FUNCTION_BLOCK FB_Tank_Target EXTENDS FB_SFC_Cycle IMPLEMENTS ITF_FB_SFC_Cycle
VAR_INPUT
	//eElementID			: E_Element_List;
	valOutlet		: E_Pis_Name;
	valLine			: E_Pis_Name;
	valTriBlender	: E_Pis_Name;
	valDrain		: E_Pis_Name;	
	valCIP			: E_Pis_Name;	
END_VAR
VAR_OUTPUT
END_VAR
VAR
	//refElement		: REFERENCE TO FB_Element;
	//refState_Long		: REFERENCE TO E_Element_State_Long;
	eReq				: E_Tank_Target;
	eProcess			: E_Tank_Target;
	eStatus				: E_Tank_Target;
	
	fbPis				: FB_Piston;
	stPis_Outlet		: REFERENCE TO ST_Piston;
	stPis_Line			: REFERENCE TO ST_Piston;
	stPis_TriBlender	: REFERENCE TO ST_Piston;
	stPis_Drain			: REFERENCE TO ST_Piston;
	stPis_CIP			: REFERENCE TO ST_Piston;

	tonDrainTime: TON;
	rt_Req_Reset: R_TRIG;
	stTankLevel			:	ST_Tank_Level	;
END_VAR
VAR_IN_OUT


END_VAR

act_GetReference();

act_Oper();
IF NOT Init.x THEN;
	act_Status();
END_IF

tonDrainTime(PT:=T#1M, 
	IN:=(eStatus=E_Tank_Target.eDrain AND stTankLevel.e_state=E_Tank_Level.eEmpty)
			OR 
		eStatus=E_Tank_Target.eClose_DrainPipe);
IF tonDrainTime.Q 
AND eReq=E_Tank_Target.eNone
AND eProcess=E_Tank_Target.eNone
THEN;
	eReq:=E_Tank_Target.eClose;
END_IF

m_Request_Reset(memo:=rt_Req_Reset);//

ACTION _aCIP_active:
bStepDone:=FALSE;
IF TRUE 
AND eStatus=E_Tank_Target.eCIP
THEN;
	bStepDone:=TRUE;
END_IF
END_ACTION

ACTION _aCIP_entry:
fbPis.m_SetByRecipe(stPis:=stPis_Outlet, 		req:=E_Piston_Recipe_State.Act);
fbPis.m_SetByRecipe(stPis:=stPis_Line, 		req:=E_Piston_Recipe_State.Release);
fbPis.m_SetByRecipe(stPis:=stPis_TriBlender, 	req:=E_Piston_Recipe_State.Release);
fbPis.m_SetByRecipe(stPis:=stPis_Drain, 		req:=E_Piston_Recipe_State.Act);
fbPis.m_SetByRecipe(stPis:=stPis_CIP, 			req:=E_Piston_Recipe_State.Act);
END_ACTION

ACTION _aClose_active:
bStepDone:=FALSE;
IF TRUE 
AND eStatus=E_Tank_Target.eClose
THEN;
	bStepDone:=TRUE;
END_IF
END_ACTION

ACTION _aClose_entry:
fbPis.m_SetByRecipe(stPis:=stPis_Outlet, 		req:=E_Piston_Recipe_State.Release);
fbPis.m_SetByRecipe(stPis:=stPis_Line, 			req:=E_Piston_Recipe_State.Release);
fbPis.m_SetByRecipe(stPis:=stPis_TriBlender, 	req:=E_Piston_Recipe_State.Release);
fbPis.m_SetByRecipe(stPis:=stPis_Drain, 		req:=E_Piston_Recipe_State.Release);
fbPis.m_SetByRecipe(stPis:=stPis_CIP, 			req:=E_Piston_Recipe_State.Release);
END_ACTION

ACTION _aDone_entry:
eProcess:=E_Tank_Target.eNone;
eReq:=E_Tank_Target.eNone;
eStatus:=E_Tank_Target.eNone;
bRun:=FALSE;
bDone:=TRUE;
END_ACTION

ACTION _aDrain_active:
bStepDone:=FALSE;
IF TRUE 
AND eStatus=E_Tank_Target.eDrain
THEN;
	bStepDone:=TRUE;
END_IF
END_ACTION

ACTION _aDrain_entry:
fbPis.m_SetByRecipe(stPis:=stPis_Outlet, 		req:=E_Piston_Recipe_State.Act);
fbPis.m_SetByRecipe(stPis:=stPis_Line, 			req:=E_Piston_Recipe_State.Release);
fbPis.m_SetByRecipe(stPis:=stPis_TriBlender, 	req:=E_Piston_Recipe_State.Release);
fbPis.m_SetByRecipe(stPis:=stPis_Drain, 		req:=E_Piston_Recipe_State.Act);
fbPis.m_SetByRecipe(stPis:=stPis_CIP, 			req:=E_Piston_Recipe_State.Release);
END_ACTION

ACTION _aDrainPipe_active:
bStepDone:=FALSE;
IF TRUE 
AND eStatus=E_Tank_Target.eClose_DrainPipe
THEN;
	bStepDone:=TRUE;
END_IF
END_ACTION

ACTION _aDrainPipe_entry:
fbPis.m_SetByRecipe(stPis:=stPis_Outlet, 		req:=E_Piston_Recipe_State.Release);
fbPis.m_SetByRecipe(stPis:=stPis_Line, 			req:=E_Piston_Recipe_State.Release);
fbPis.m_SetByRecipe(stPis:=stPis_TriBlender, 	req:=E_Piston_Recipe_State.Release);
fbPis.m_SetByRecipe(stPis:=stPis_Drain, 		req:=E_Piston_Recipe_State.Act);
fbPis.m_SetByRecipe(stPis:=stPis_CIP, 			req:=E_Piston_Recipe_State.Release);
END_ACTION

ACTION _aInit_active:
SFCReset:=FALSE;
END_ACTION

ACTION _aInit_exit:
eProcess:=E_Tank_Target.eNone;
eReq:=E_Tank_Target.eNone;
END_ACTION

ACTION _aOpen_active:
bStepDone:=FALSE;
IF TRUE 
AND eStatus=E_Tank_Target.eOpen
THEN;
	bStepDone:=TRUE;
END_IF
END_ACTION

ACTION _aOpen_entry:
fbPis.m_SetByRecipe(stPis:=stPis_Outlet, req:=E_Piston_Recipe_State.Act);
//fbPis.m_SetByRecipe(stPis:=valLine, req:=E_Piston_Recipe_State.Release);
//fbPis.m_SetByRecipe(stPis:=valTriBlender, req:=E_Piston_Recipe_State.Release);
fbPis.m_SetByRecipe(stPis:=stPis_Drain, req:=E_Piston_Recipe_State.Release);
fbPis.m_SetByRecipe(stPis:=stPis_CIP, req:=E_Piston_Recipe_State.Release);
END_ACTION

ACTION _aReady_active:

eStatus:=E_Tank_Target.eNone;
CASE eReq OF
	E_Tank_Target.eClose:;
			IF TRUE THEN;
				eProcess:=E_Tank_Target.eClose;
			END_IF

	E_Tank_Target.eOpen:;
			IF TRUE THEN;
				eProcess:=E_Tank_Target.eOpen;
			END_IF	
			
	E_Tank_Target.eDrain:;
			IF TRUE THEN;
				eProcess:=E_Tank_Target.eDrain;
			END_IF
	
	E_Tank_Target.eClose_DrainPipe:;
			IF TRUE THEN;
				eProcess:=E_Tank_Target.eClose_DrainPipe;
			END_IF	
			
	E_Tank_Target.eCIP:;
			IF TRUE THEN;
				eProcess:=E_Tank_Target.eCIP;
			END_IF	

END_CASE
END_ACTION

ACTION _aReady_exit:
bRun:=TRUE;
bDone:=FALSE;
END_ACTION

ACTION act_GetReference:
m_Set_SFCFlags_Reference();
//refElement REF= fbElement[eElementID];
//refState_Long REF= fbElement[eElementID].eState_Long;

stPis_Outlet		REF= g_Piston.stPis[valOutlet];
stPis_Line			REF= g_Piston.stPis[valLine];
stPis_TriBlender	REF= g_Piston.stPis[valTriBlender];
stPis_Drain			REF= g_Piston.stPis[valDrain];
stPis_CIP			REF= g_Piston.stPis[valCIP];
END_ACTION

ACTION act_Oper:
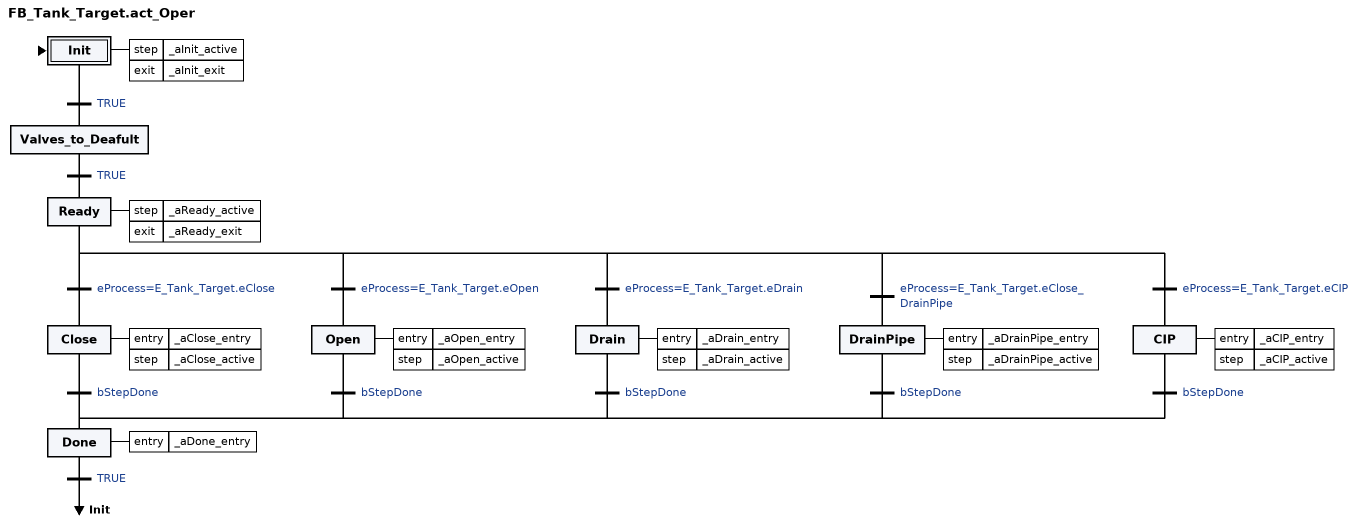
INITIAL_STEP Init:  // min time T#0.5s
    _aInit_active(N);  // step action
    _aInit_exit(P0);  // exit action
END_STEP
TRANSITION FROM Init TO Valves_to_Deafult
    := TRUE;
END_TRANSITION
STEP Valves_to_Deafult:
END_STEP
TRANSITION FROM Valves_to_Deafult TO Ready
    := TRUE;
END_TRANSITION
STEP Ready:
    _aReady_active(N);  // step action
    _aReady_exit(P0);  // exit action
END_STEP
TRANSITION FROM Ready TO Close
    := eProcess=E_Tank_Target.eClose;
END_TRANSITION
STEP Close:
    _aClose_entry(P1);  // entry action
    _aClose_active(N);  // step action
END_STEP
TRANSITION FROM Close TO Done
    := bStepDone;
END_TRANSITION
TRANSITION FROM Ready TO Open
    := eProcess=E_Tank_Target.eOpen;
END_TRANSITION
STEP Open:
    _aOpen_entry(P1);  // entry action
    _aOpen_active(N);  // step action
END_STEP
TRANSITION FROM Open TO Done
    := bStepDone;
END_TRANSITION
TRANSITION FROM Ready TO Drain
    := eProcess=E_Tank_Target.eDrain;
END_TRANSITION
STEP Drain:
    _aDrain_entry(P1);  // entry action
    _aDrain_active(N);  // step action
END_STEP
TRANSITION FROM Drain TO Done
    := bStepDone;
END_TRANSITION
TRANSITION FROM Ready TO DrainPipe
    := eProcess=E_Tank_Target.eClose_DrainPipe;
END_TRANSITION
STEP DrainPipe:
    _aDrainPipe_entry(P1);  // entry action
    _aDrainPipe_active(N);  // step action
END_STEP
TRANSITION FROM DrainPipe TO Done
    := bStepDone;
END_TRANSITION
TRANSITION FROM Ready TO CIP
    := eProcess=E_Tank_Target.eCIP;
END_TRANSITION
STEP CIP:
    _aCIP_entry(P1);  // entry action
    _aCIP_active(N);  // step action
END_STEP
TRANSITION FROM CIP TO Done
    := bStepDone;
END_TRANSITION
STEP Done:  // min time T#0.2s
    _aDone_entry(P1);  // entry action
END_STEP
TRANSITION FROM Done TO Init
    := TRUE;
END_TRANSITION
// branch label Branch0_act_Oper_Tank
END_ACTION

ACTION act_Status:


IF TRUE 
AND fbPis.m_CheckByRecipe(stPis:=stPis_Outlet, 		req:=E_Piston_Recipe_State.Release)
AND fbPis.m_CheckByRecipe(stPis:=stPis_Line, 		req:=E_Piston_Recipe_State.Release)
AND fbPis.m_CheckByRecipe(stPis:=stPis_TriBlender, 	req:=E_Piston_Recipe_State.Release)
AND fbPis.m_CheckByRecipe(stPis:=stPis_Drain, 		req:=E_Piston_Recipe_State.Release)
AND fbPis.m_CheckByRecipe(stPis:=stPis_CIP, 		req:=E_Piston_Recipe_State.Release)
THEN;
	eStatus:=E_Tank_Target.eClose;
	
ELSIF TRUE 
AND fbPis.m_CheckByRecipe(stPis:=stPis_Outlet, 		req:=E_Piston_Recipe_State.Act)
//AND fbPis.m_CheckByRecipe(stPis:=valLine, 		req:=E_Piston_Recipe_State.Release)
//AND fbPis.m_CheckByRecipe(stPis:=valTriBlender, 	req:=E_Piston_Recipe_State.Release)
AND fbPis.m_CheckByRecipe(stPis:=stPis_Drain, 		req:=E_Piston_Recipe_State.Release)
AND fbPis.m_CheckByRecipe(stPis:=stPis_CIP, 		req:=E_Piston_Recipe_State.Release)
THEN;
	eStatus:=E_Tank_Target.eOpen;
	
ELSIF TRUE 
AND fbPis.m_CheckByRecipe(stPis:=stPis_Outlet, 		req:=E_Piston_Recipe_State.Act)
AND fbPis.m_CheckByRecipe(stPis:=stPis_Line, 		req:=E_Piston_Recipe_State.Release)
AND fbPis.m_CheckByRecipe(stPis:=stPis_TriBlender, 	req:=E_Piston_Recipe_State.Release)
AND fbPis.m_CheckByRecipe(stPis:=stPis_Drain, 		req:=E_Piston_Recipe_State.Act)
AND fbPis.m_CheckByRecipe(stPis:=stPis_CIP, 		req:=E_Piston_Recipe_State.Release)
THEN;
	eStatus:=E_Tank_Target.eDrain;
	
ELSIF TRUE 
AND fbPis.m_CheckByRecipe(stPis:=stPis_Outlet, 		req:=E_Piston_Recipe_State.Release)
AND fbPis.m_CheckByRecipe(stPis:=stPis_Line, 		req:=E_Piston_Recipe_State.Release)
AND fbPis.m_CheckByRecipe(stPis:=stPis_TriBlender, 	req:=E_Piston_Recipe_State.Release)
AND fbPis.m_CheckByRecipe(stPis:=stPis_Drain, 		req:=E_Piston_Recipe_State.Act)
AND fbPis.m_CheckByRecipe(stPis:=stPis_CIP, 		req:=E_Piston_Recipe_State.Release)
THEN;
	eStatus:=E_Tank_Target.eClose_DrainPipe;
	
ELSIF TRUE 
AND fbPis.m_CheckByRecipe(stPis:=stPis_Outlet, 		req:=E_Piston_Recipe_State.Act)
AND fbPis.m_CheckByRecipe(stPis:=stPis_Line, 		req:=E_Piston_Recipe_State.Release)
AND fbPis.m_CheckByRecipe(stPis:=stPis_TriBlender, 	req:=E_Piston_Recipe_State.Release)
AND fbPis.m_CheckByRecipe(stPis:=stPis_Drain, 		req:=E_Piston_Recipe_State.Act)
AND fbPis.m_CheckByRecipe(stPis:=stPis_CIP, 		req:=E_Piston_Recipe_State.Act)
THEN;
	eStatus:=E_Tank_Target.eCIP;
	
ELSE;
	eStatus:=E_Tank_Target.eNone;
END_IF
END_ACTION

METHOD m_CheckStatus : BOOL
VAR_INPUT
	eReqStatus		: E_Tank_Target;
END_VAR
IF eStatus=eReqStatus 
AND eProcess=E_Tank_Target.eNone
AND eReq=E_Tank_Target.eNone
AND bReady
AND bDone
AND NOT bRun
THEN;
	m_CheckStatus:=TRUE;
END_IF
END_METHOD

METHOD m_Request_Reset : BOOL
VAR_IN_OUT
	memo: R_TRIG;
END_VAR
memo(CLK:=eReq=0);
IF TRUE 
AND memo.Q
THEN;
	SFCReset:=TRUE;
END_IF
END_METHOD

METHOD m_Run : BOOL
VAR_INPUT
	eReqProc			: E_Tank_Target;
END_VAR
IF eProcess=E_Tank_Target.eNone THEN;
	eProcess:=eReq:=eReqProc;
	bDone:=FALSE;
	m_Run:=TRUE;
END_IF
END_METHOD

METHOD m_Set_SFCFlags_Reference : BOOL
//Set reference to SFC flags

refSFC.SFCInit REF= SFCInit;
refSFC.SFCReset REF= SFCReset;
refSFC.SFCError REF= SFCError;
refSFC.SFCEnableLimit REF= SFCEnableLimit;
refSFC.SFCErrorStep REF= SFCErrorStep;
refSFC.SFCErrorPOU REF= SFCErrorPOU;
refSFC.SFCQuitError REF= SFCQuitError;
refSFC.SFCPause REF= SFCPause;
refSFC.SFCTrans REF= SFCTrans;
refSFC.SFCCurrentStep REF= SFCCurrentStep;
refSFC.SFCTip REF= SFCTip;
refSFC.SFCTipMode REF= SFCTipMode;

// Cycle handle for SFC
m_SFC_Handle();
END_METHOD

METHOD set_TankLevel : BOOL
VAR_INPUT
	set_stTankLevel			:	ST_Tank_Level	;
END_VAR
stTankLevel:=set_stTankLevel;
END_METHOD

END_FUNCTION_BLOCK

(* stored: Version 1.1.0.1, ProductVersion 3.1.4024.13
   POU FB_Tank_Target: Id {e77bc243-ef67-4877-849d-f4a841448420}, SpecialFunc None
   Folder Manage: Id {e461fcff-545d-4d57-a27d-4174ff6e3a51}
   Action _aCIP_active: Id {e16ca9a6-461a-481e-961d-0ed26f76e308}
   Action _aCIP_entry: Id {a141e873-c7fc-4307-9c91-bb51c75dad2b}
   Action _aClose_active: Id {d079a344-74ba-42ce-88cf-aed803eb2b19}
   Action _aClose_entry: Id {db19abbe-579c-4574-a1a2-48f247faffd5}
   Action _aDone_entry: Id {1342fd33-e78f-4125-a323-9d65d6a85b09}
   Action _aDrain_active: Id {f02cc56e-f572-40d0-ba02-338281ca63e4}
   Action _aDrain_entry: Id {59a8b0e3-9d73-4126-9788-a378683e6b96}
   Action _aDrainPipe_active: Id {0a536e01-1fe5-4e37-aa4a-59dcbfe014c1}
   Action _aDrainPipe_entry: Id {70d2d20b-108b-48e4-bd4d-c6eb6f3e46be}
   Action _aInit_active: Id {cef529ac-1147-479f-874c-293fab5d64a2}
   Action _aInit_exit: Id {883cd8f7-e2c9-4fd3-a843-28ad6c843fc3}
   Action _aOpen_active: Id {091a9747-c4fd-474e-986a-8d9d28db4c2e}
   Action _aOpen_entry: Id {40cbadc0-1a08-4490-ae58-09b056231ca7}
   Action _aReady_active: Id {11ea1fd0-5021-4a91-99b3-72574a941116}
   Action _aReady_exit: Id {10d9b54d-9a6f-4993-86ba-c8a5bc0d174a}
   Action act_GetReference: Id {cf9432c7-1e36-4aaf-9faf-4cb2c932a09a}
   Action act_Oper: Id {62af6f6a-742c-430d-9588-934f1d656471}
   Action act_Status: Id {0d6b2513-8aec-4f27-b7af-4e0f232d3f1f}
   Method m_CheckStatus: Id {730e0eab-fcbe-441f-8132-795becd278a2}
   Method m_Request_Reset: Id {06b07d97-a5cd-434a-8128-1378a573a1f8}
   Method m_Run: Id {7ffc4675-e14a-4e0d-a035-300d182aa227}
   Method m_Set_SFCFlags_Reference: Id {f4d4034f-fbcd-4ba0-9568-d6c2136b33ee}
   Method set_TankLevel: Id {2976f91a-4f21-42e1-852d-f74c3c86612b} *)
